Fanuc KAREL source: kt00302.KL

-- PROVISIONAL review KL for V1013-1; original PC SHA256 93e4615c5a4b092bd1b063ab247f0e8c9188fb1d7dfb9a491f40a172e73db85c
-- Incomplete behavior may be omitted. Consult companion uncertainty JSON. Do not deploy.
PROGRAM KT00302
%NOLOCKGROUP
VAR
  S1 : STRING[80]
  S2 : STRING[80]
  OUT : BOOLEAN
BEGIN
  -- UNRESOLVED_PC offsets 5-14; opcodes 3F,75
  -- UNRESOLVED_PC offsets 19-28; opcodes 3F,75
  -- UNRESOLVED_PC offsets 33-42; opcodes 3F,75
  -- UNRESOLVED_PC offsets 47-56; opcodes 3F,75
  -- UNRESOLVED_PC offsets 61-80; opcodes 73,73,84,23
  -- UNRESOLVED_PC offsets 85-89; opcodes 7F
END KT00302
